Fanuc KAREL source: kt00869.KL

-- PROVISIONAL review KL for V940-1; original PC SHA256 47eba381261ba0f90bfa3d82c6dea36029eda366b20c83dee3d34a7dcc88c95f
-- Incomplete behavior may be omitted. Consult companion uncertainty JSON. Do not deploy.
PROGRAM KT00869
%NOLOCKGROUP
VAR
  I1 : INTEGER
  I2 : INTEGER
  OUT : REAL
BEGIN
  -- V9_ZERO_TABLE_METADATA_HINT layout=0001; no indexed target words; source/name/runtime held
  -- UNRESOLVED_PC offsets 5-16; opcodes 2E,23
  -- UNRESOLVED_PC offsets 21-32; opcodes 2E,23
  -- UNRESOLVED_PC offsets 37-48; opcodes 2E,23
  -- UNRESOLVED_PC offsets 53-64; opcodes 2E,23
  -- UNRESOLVED_PC offsets 69-87; opcodes 27,27,21,64,76,64,23
  -- UNRESOLVED_PC offsets 92-96; opcodes 7F
END KT00869
